(* IEC 61131-3 sources: codesys-framework/txt/application/WeVe Core (library)/50 Component/FB_Component, 6 files *)

(* ---- Busy.prop.st ---- *)
PROPERTY Busy : BOOL

// --- BEGIN IMPLEMENTATION ---

// ----------- GET -----------
VAR
END_VAR

// -- BEGIN IMPLEMENTATION GET --
Busy := _xBusy;

(* ---- Done.prop.st ---- *)
PROPERTY Done : BOOL

// --- BEGIN IMPLEMENTATION ---

// ----------- GET -----------
VAR
END_VAR

// -- BEGIN IMPLEMENTATION GET --
Done := _xDone;

(* ---- Error.prop.st ---- *)
{attribute 'monitoring' := 'variable'}
PROPERTY Error : SC_Error
// --- BEGIN IMPLEMENTATION ---

// ----------- GET -----------
VAR
END_VAR

// -- BEGIN IMPLEMENTATION GET --
Error := _scError;

(* ---- Initialize.method.st ---- *)
METHOD Initialize
VAR_INPUT
END_VAR

// --- BEGIN IMPLEMENTATION ---

_xBusy := FALSE;
_xDone := FALSE;

(* ---- Name.prop.st ---- *)
PROPERTY Name : STRING
// --- BEGIN IMPLEMENTATION ---

// ----------- GET -----------
VAR
END_VAR

// -- BEGIN IMPLEMENTATION GET --
Name := _sName;

// ----------- SET -----------
PUBLIC
VAR
END_VAR

// -- BEGIN IMPLEMENTATION SET --
_sName := Name;

(* ---- Reset.method.st ---- *)
METHOD Reset : BOOL
VAR_INPUT
END_VAR

// --- BEGIN IMPLEMENTATION ---

_scError.xErrorActive := FALSE;
_scError.sError := '';
